FUNCTION_BLOCK fbMonoSwitch IMPLEMENTS iSwitch
VAR
	Input AT %I* : BOOL;					// Physical switch input
	
	SwitchPressed : R_TRIG;
	SwitchReleased : F_Trig;
END_VAR

SwitchPressed(CLK := Input);
SwitchReleased(CLK := Input);

PROPERTY PUBLIC IsPressed : BOOL
GET
IsPressed := SwitchPressed.Q;
END_GET
END_PROPERTY

PROPERTY IsReleased : BOOL
GET
IsReleased := SwitchReleased.Q;
END_GET
END_PROPERTY

END_FUNCTION_BLOCK

(* stored: Version 1.1.0.1
   POU fbMonoSwitch: Id {21737aef-df48-4987-83e0-aae9b7cbc7ab}, SpecialFunc None
   Property IsPressed: Id {238fedb4-7f31-449e-bffb-88405f0e3fe6}
   Get Get: Id {bc4b2b4d-b425-4031-ada5-782516be3c69}
   Property IsReleased: Id {f2e12f74-1423-4b11-9d68-63053027c6bb}
   Get Get: Id {00b0c95b-d4ed-4500-978f-f246b06ade20} *)
